// Mitsubishi GX Works2 project: IAN - SOCKET MODBUSTCP   PLC: Q03UDV

PROGRAM MAIN
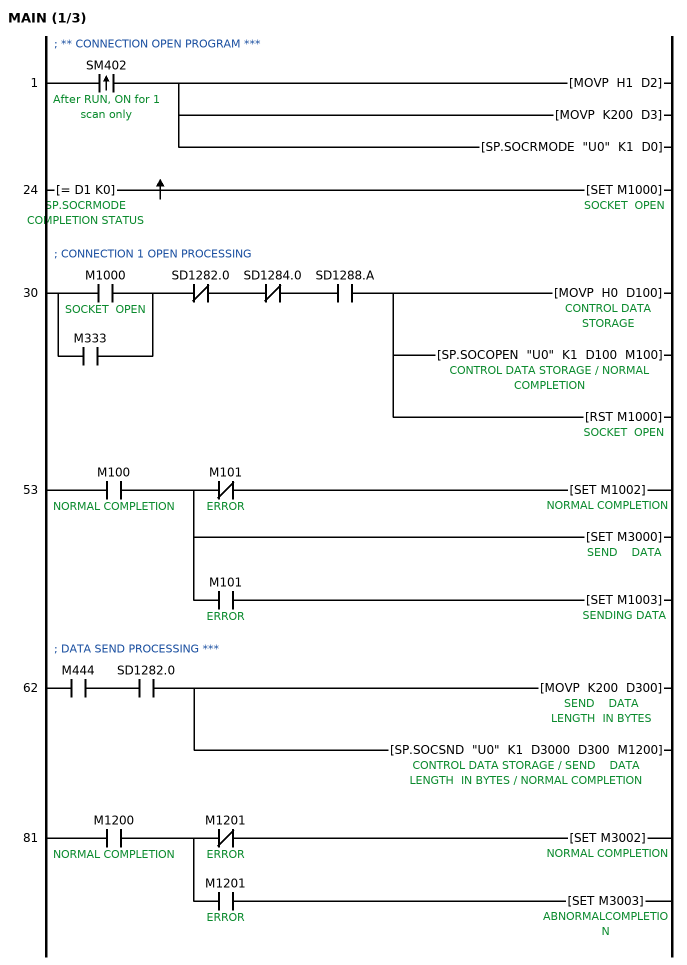
; ** CONNECTION OPEN PROGRAM ***
1     LDP     SM402  ; After RUN, ON for 1 scan only
      MOVP    H1 D2
        [note] TCP RECEIVE MODE (SET TO VAR)
      MOVP    K200 D3
        [note] RECEIVE DATA SIZE IN BYTES
      SP.SOCRMODE "U0" K1 D0
        [note] CON. 1 TCP RECEIVE MODE CHANGE
24    LD=     D1 K0  ; SP.SOCRMODE COMPLETION STATUS
      MEP
      SET     M1000  ; SOCKET  OPEN
; CONNECTION 1 OPEN PROCESSING
30    LD      M1000  ; SOCKET  OPEN
      OR      M333
      ANI     SD1282.0
      ANI     SD1284.0
      AND     SD1288.A
      MOVP    H0 D100  ; CONTROL DATA STORAGE
        [note] EXECUTION/COMPLETION TYPE
      SP.SOCOPEN "U0" K1 D100 M100  ; NORMAL COMPLETION
      RST     M1000  ; SOCKET  OPEN
53    LD      M100  ; NORMAL COMPLETION
      MPS
      ANI     M101  ; ERROR
      SET     M1002  ; NORMAL COMPLETION
      MPP
      SET     M3000  ; SEND    DATA
      AND     M101  ; ERROR
      SET     M1003  ; SENDING DATA
; DATA SEND PROCESSING ***
62    LD      M444
      AND     SD1282.0
      MOVP    K200 D300  ; SEND    DATA    LENGTH  IN BYTES
        [note] SEND DATA LENGTH
      SP.SOCSND "U0" K1 D3000 D300 M1200  ; CONTROL DATA STORAGE / NORMAL COMPLETION
81    LD      M1200  ; NORMAL COMPLETION
      MPS
      ANI     M1201  ; ERROR
      SET     M3002  ; NORMAL COMPLETION
      MPP
      AND     M1201  ; ERROR
      SET     M3003  ; ABNORMALCOMPLETION
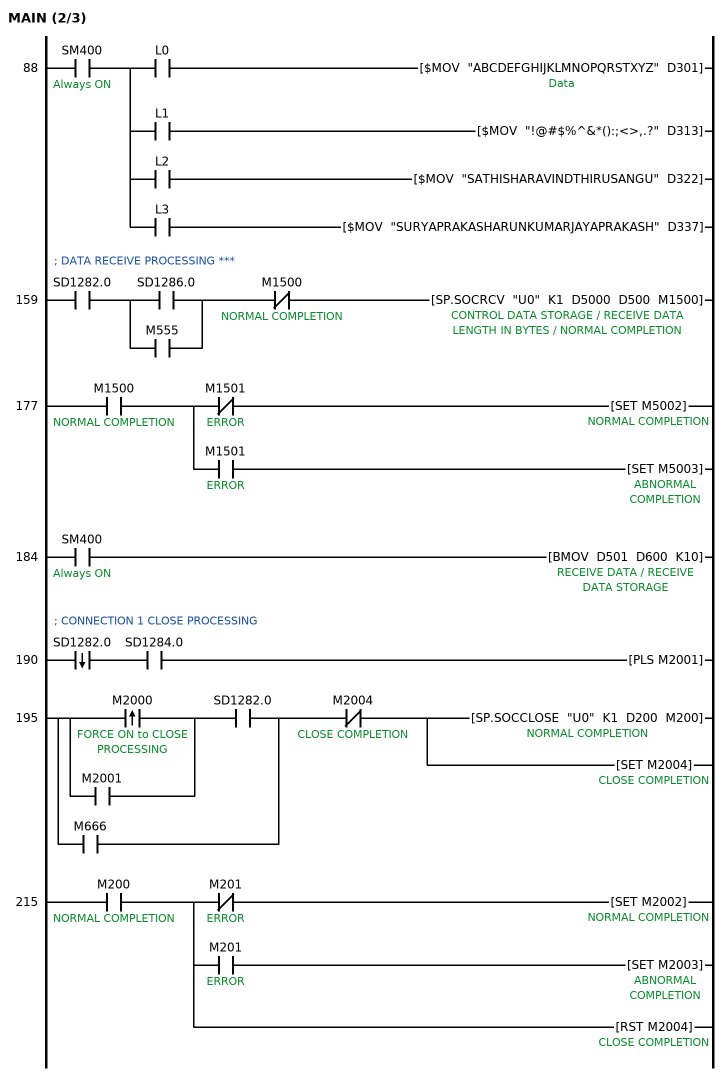
88    LD      SM400  ; Always ON
      MPS
      AND     L0
      $MOV    "ABCDEFGHIJKLMNOPQRSTXYZ" D301  ; Data
      MRD
      AND     L1
      $MOV    "!@#$%^&*():;<>,.?" D313
      MRD
      AND     L2
      $MOV    "SATHISHARAVINDTHIRUSANGU" D322
      MPP
      AND     L3
      $MOV    "SURYAPRAKASHARUNKUMARJAYAPRAKASH" D337
; DATA RECEIVE PROCESSING ***
159   LD      SD1282.0
      LD      SD1286.0
      OR      M555
      ANB
      ANI     M1500  ; NORMAL COMPLETION
      SP.SOCRCV "U0" K1 D5000 D500 M1500  ; CONTROL DATA STORAGE / RECEIVE DATA LENGTH IN BYTES
177   LD      M1500  ; NORMAL COMPLETION
      MPS
      ANI     M1501  ; ERROR
      SET     M5002  ; NORMAL COMPLETION
      MPP
      AND     M1501  ; ERROR
      SET     M5003  ; ABNORMAL COMPLETION
184   LD      SM400  ; Always ON
      BMOV    D501 D600 K10  ; RECEIVE DATA / RECEIVE DATA STORAGE
; CONNECTION 1 CLOSE PROCESSING
190   LDF     SD1282.0
      AND     SD1284.0
      PLS     M2001
195   LDP     M2000  ; FORCE ON to CLOSE PROCESSING
      OR      M2001
      AND     SD1282.0
      OR      M666
      ANI     M2004  ; CLOSE COMPLETION
      SP.SOCCLOSE "U0" K1 D200 M200  ; NORMAL COMPLETION
      SET     M2004  ; CLOSE COMPLETION
215   LD      M200  ; NORMAL COMPLETION
      MPS
      ANI     M201  ; ERROR
      SET     M2002  ; NORMAL COMPLETION
      MRD
      AND     M201  ; ERROR
      SET     M2003  ; ABNORMAL COMPLETION
      MPP
      RST     M2004  ; CLOSE COMPLETION
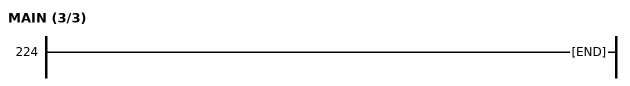
224   END
END_PROGRAM

// device comments not shown above
M1050  ; SOCKET OPEN
M1053  ; ABNORMAL
M1150  ; SOCKET OPEN
M1153  ; ABNORMAL
M3050  ; SEND    DATA
M3150  ; SEND DATA
M5103  ; ABNORMAL COMPLETION
M5203  ; ABNORMAL COMPLETION
D550  ; RECEIVE VALUE 567 from 2nd SLAVE
D610  ; RECEIVE VALUE 234 from 1st SLAVE
D620  ; RECEIVE VALUE 567 from 2nd SLAVE
D630  ; RECEIVE VALUE 789 from 3rd SLAVE
D1600  ; SEND    DATA    LENGTH  IN BYTES
D1601  ; SENDING 123 to 2nd STATION D500
D1700  ; SEND    DATA    LENGTH  IN BYTES
D1701  ; SENDING 123 to 3rd STATION D500
